TYPE stLightCmdEvent :
STRUCT
	Execute : BOOL;
	TargetState : stLightState;
	Source  : eLightCmdSource;
END_STRUCT
END_TYPE

(* stored: Version 1.1.0.1
   DUT stLightCmdEvent: Id {b3ebb80a-5323-4b41-8ea8-2a1f2cbf09f2} *)
